(* IEC 61131-3 sources: llm-plc-st-eval/data/processed_definitivo/claude-sonnet-4-6/A3/few_shot, 3 files *)

(* ---- ejec_1.st ---- *)
FUNCTION_BLOCK FB_Com
VAR_INPUT
    txReq  : BOOL; (* Solicitud de inicio de intercambio *)
    rxOk   : BOOL; (* Confirmacion de recepcion del dispositivo externo *)
    rxData : INT;  (* Dato recibido del dispositivo externo *)
END_VAR
VAR_OUTPUT
    txData   : INT;  (* Dato transmitido al dispositivo externo *)
    ocupado  : BOOL; (* Intercambio en curso *)
    ok       : BOOL; (* Intercambio completado con exito *)
    error    : BOOL; (* Fallaron los 3 intentos *)
    nIntentos: INT;  (* Numero del intento en curso o ultimo realizado *)
END_VAR
VAR
    tIntento   : TON;        (* Temporizador de plazo por intento: 500 ms *)
    txReq_prev : BOOL;       (* Valor anterior de txReq para detectar flanco *)
    flanco     : BOOL;       (* Flanco ascendente de txReq *)
    rxOk_prev  : BOOL;       (* Valor anterior de rxOk para detectar flanco *)
    flancoRx   : BOOL;       (* Flanco ascendente de rxOk *)
    TX_VALUE   : INT := 100; (* Valor de prueba fijo a transmitir *)
    MAX_INT    : INT := 3;   (* Numero maximo de intentos *)
END_VAR

(* --- Deteccion de flancos ascendentes --- *)
flanco   := txReq  AND NOT txReq_prev;
flancoRx := rxOk   AND NOT rxOk_prev;

(* --- Inicio de un nuevo intercambio (solo si no hay uno en curso) --- *)
IF flanco AND NOT ocupado THEN
    ocupado   := TRUE;
    ok        := FALSE;
    error     := FALSE;
    nIntentos := 1;
    txData    := TX_VALUE;
    tIntento(IN := FALSE, PT := T#500MS); (* Reset del temporizador *)
END_IF;

(* --- Logica principal durante un intercambio en curso --- *)
IF ocupado THEN
    (* Arrancar/mantener el temporizador del intento actual *)
    tIntento(IN := TRUE, PT := T#500MS);

    (* Caso 1: respuesta correcta dentro del plazo *)
    IF flancoRx AND (rxData = TX_VALUE) AND NOT tIntento.Q THEN
        ocupado  := FALSE;
        ok       := TRUE;
        tIntento(IN := FALSE, PT := T#500MS); (* Detener temporizador *)

    (* Caso 2: plazo vencido sin confirmacion, o respuesta con dato incorrecto *)
    ELSIF tIntento.Q OR (flancoRx AND (rxData <> TX_VALUE)) THEN
        IF nIntentos < MAX_INT THEN
            (* Iniciar siguiente intento *)
            nIntentos := nIntentos + 1;
            tIntento(IN := FALSE, PT := T#500MS); (* Reset para nuevo plazo *)
        ELSE
            (* Se agotaron los 3 intentos *)
            ocupado := FALSE;
            error   := TRUE;
            tIntento(IN := FALSE, PT := T#500MS); (* Detener temporizador *)
        END_IF;
    END_IF;
END_IF;

(* --- Guardar estados anteriores para proxima ejecucion --- *)
txReq_prev := txReq;
rxOk_prev  := rxOk;

END_FUNCTION_BLOCK

(* ---- ejec_2.st ---- *)
FUNCTION_BLOCK FB_Com
VAR_INPUT
    txReq  : BOOL; (* Solicitud de inicio de intercambio *)
    rxOk   : BOOL; (* Confirmacion recibida del dispositivo externo *)
    rxData : INT;  (* Dato recibido (eco esperado) *)
END_VAR
VAR_OUTPUT
    txData   : INT;  (* Dato transmitido al dispositivo externo *)
    ocupado  : BOOL; (* TRUE mientras hay un intercambio en curso *)
    ok       : BOOL; (* TRUE si el intercambio termino correctamente *)
    error    : BOOL; (* TRUE si fallaron los 3 intentos *)
    nIntentos: INT;  (* Numero del intento en curso o ultimo realizado *)
END_VAR
VAR
    tIntento  : TON;       (* Temporizador de plazo por intento (500 ms) *)
    txReqPrev : BOOL;      (* Valor anterior de txReq para detectar flanco *)
    enCurso   : BOOL;      (* Intercambio activo internamente *)
    VAL_PRUEBA: INT := 100;(* Valor fijo de prueba transmitido *)
END_VAR

(* --- Deteccion de flanco ascendente en txReq --- *)
IF txReq AND NOT txReqPrev THEN
    IF NOT enCurso THEN
        (* Iniciar nuevo intercambio *)
        enCurso   := TRUE;
        ocupado   := TRUE;
        ok        := FALSE;
        error     := FALSE;
        nIntentos := 1;
        txData    := VAL_PRUEBA;
        (* Arrancar temporizador del primer intento *)
        tIntento(IN := FALSE, PT := T#500MS); (* Reset previo *)
    END_IF;
END_IF;
txReqPrev := txReq;

(* --- Logica principal del intercambio --- *)
IF enCurso THEN
    (* Mantener temporizador activo *)
    tIntento(IN := TRUE, PT := T#500MS);

    (* Comprobar respuesta correcta: rxOk activo y eco coincide *)
    IF rxOk AND (rxData = txData) THEN
        (* Intento exitoso *)
        ok        := TRUE;
        ocupado   := FALSE;
        enCurso   := FALSE;
        tIntento(IN := FALSE, PT := T#500MS); (* Detener temporizador *)

    (* Comprobar fallo: plazo vencido O rxOk con dato incorrecto *)
    ELSIF tIntento.Q OR (rxOk AND (rxData <> txData)) THEN
        (* Detener temporizador antes de evaluar siguiente paso *)
        tIntento(IN := FALSE, PT := T#500MS);

        IF nIntentos >= 3 THEN
            (* Agotados los 3 intentos *)
            error   := TRUE;
            ocupado := FALSE;
            enCurso := FALSE;
        ELSE
            (* Iniciar siguiente intento *)
            nIntentos := nIntentos + 1;
            (* El temporizador se reanudara en el proximo ciclo con IN=TRUE *)
        END_IF;
    END_IF;
END_IF;

END_FUNCTION_BLOCK

(* ---- ejec_3.st ---- *)
FUNCTION_BLOCK FB_Com
VAR_INPUT
    txReq  : BOOL; (* Solicitud de inicio de intercambio *)
    rxOk   : BOOL; (* Confirmacion recibida del dispositivo externo *)
    rxData : INT;  (* Dato recibido (eco esperado) *)
END_VAR
VAR_OUTPUT
    txData   : INT;  (* Dato transmitido al dispositivo externo *)
    ocupado  : BOOL; (* Intercambio en curso *)
    ok       : BOOL; (* Ultimo intercambio exitoso *)
    error    : BOOL; (* Fallaron los 3 intentos *)
    nIntentos: INT;  (* Numero del intento en curso *)
END_VAR
VAR
    tTimeout  : TON;          (* Temporizador de plazo por intento *)
    txReqPrev : BOOL;         (* Valor anterior de txReq para detectar flanco *)
    activo    : BOOL;         (* Intercambio en curso (interno) *)
    txValor   : INT := 100;   (* Valor de prueba fijo *)
END_VAR

(* --- Deteccion de flanco ascendente en txReq --- *)
IF txReq AND NOT txReqPrev AND NOT activo THEN
    (* Inicio de nuevo intercambio *)
    activo    := TRUE;
    ocupado   := TRUE;
    ok        := FALSE;
    error     := FALSE;
    nIntentos := 1;
    txData    := txValor;
    tTimeout(IN := FALSE, PT := T#500MS); (* Reset del temporizador *)
END_IF;
txReqPrev := txReq;

(* --- Logica principal del intercambio --- *)
IF activo THEN
    (* Ejecutar temporizador del intento actual *)
    tTimeout(IN := TRUE, PT := T#500MS);

    (* Verificar respuesta correcta: rxOk activo y eco correcto *)
    IF rxOk AND (rxData = txValor) THEN
        (* Intento exitoso *)
        ok       := TRUE;
        ocupado  := FALSE;
        activo   := FALSE;
        tTimeout(IN := FALSE, PT := T#500MS); (* Detener temporizador *)

    (* Verificar fallo: plazo vencido o eco incorrecto *)
    ELSIF tTimeout.Q OR (rxOk AND (rxData <> txValor)) THEN
        tTimeout(IN := FALSE, PT := T#500MS); (* Reset del temporizador *)

        IF nIntentos < 3 THEN
            (* Iniciar siguiente intento *)
            nIntentos := nIntentos + 1;
            (* El temporizador arrancara en el proximo ciclo con IN=TRUE *)
        ELSE
            (* Agotados los 3 intentos: error *)
            error   := TRUE;
            ocupado := FALSE;
            activo  := FALSE;
        END_IF;
    END_IF;
END_IF;

END_FUNCTION_BLOCK
